FUNCTION_BLOCK AutomaticOperation (* Basic Function Block Type *)
  (* Standard: 61499-2 *)
  (* Version 0.0, 10/19/2026, macie, Schneider Electric, Template *)
  PACKAGE Main;
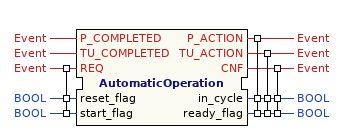
  EVENT_INPUT
    P_COMPLETED; (* Normal Execution Request *)
    TU_COMPLETED;
    REQ WITH reset_flag, start_flag;
  END_EVENT
  EVENT_OUTPUT
    P_ACTION WITH in_cycle, ready_flag; (* Execution Confirmation *)
    TU_ACTION WITH in_cycle, ready_flag;
    CNF WITH in_cycle, ready_flag;
  END_EVENT
  VAR_INPUT
    reset_flag : BOOL := FALSE;
    start_flag : BOOL := FALSE;
  END_VAR
  VAR_OUTPUT
    in_cycle : BOOL := FALSE;
    ready_flag : BOOL := TRUE;
  END_VAR
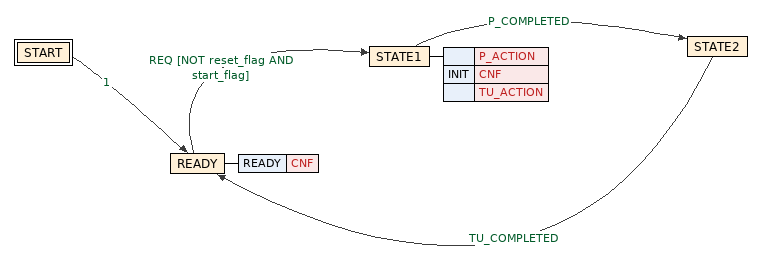
  EC_STATES
    START; (* Initial State *)
    READY : READY -> CNF;
    STATE1 : -> P_ACTION, INIT -> CNF, -> TU_ACTION;
    STATE2;
  END_STATES
  EC_TRANSITIONS
    START TO READY := 1;
    READY TO STATE1 := REQ [NOT reset_flag AND start_flag];
    STATE1 TO STATE2 := P_COMPLETED;
    STATE2 TO READY := TU_COMPLETED;
  END_TRANSITIONS
  ALGORITHM INIT IN ST: (* Initialization algorithm *)
;
ready_flag := FALSE;
in_cycle := TRUE;
  END_ALGORITHM
  ALGORITHM STEP1 IN ST: (* Normally executed algorithm *)
;
in_cycle := TRUE;
  END_ALGORITHM
  ALGORITHM STEP2 IN ST:
;
  END_ALGORITHM
  ALGORITHM STEP3 IN ST:
;
  END_ALGORITHM
  ALGORITHM STEP4 IN ST:
;
  END_ALGORITHM
  ALGORITHM STEP0 IN ST:
;

ready_flag := FALSE;
  END_ALGORITHM
  ALGORITHM READY IN ST:
;
ready_flag := TRUE;
in_cycle := FALSE;
  END_ALGORITHM
END_FUNCTION_BLOCK
